(* CODESYS project Visualization.vis.xml

Project tree, tasks and I/O mapping:
  visualisation Visualization
*)

// /Visualization
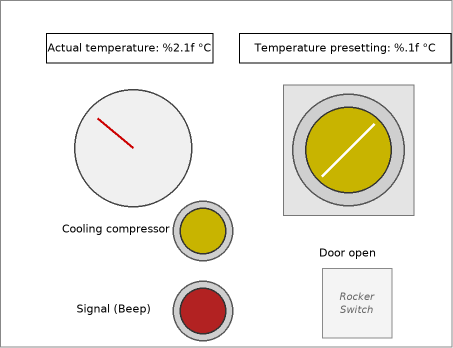
VISUALIZATION Visualization  // 453x348
    Rectangle (46,33 167x30), "Actual temperature: %2.1f °C", text variable: Glob_Var.TempActual
    Lamp1 (168,196 70x70), variable: Glob_Var.Compressor, style: Lamp-Lamp1-Yellow
    Rectangle (239,33 212x30), "Temperature presetting: %.1f °C", text variable: Glob_Var.TempSet
        OnMouseDown: write the text variable via Default, min 3, max 12
    Potentiometer360 (283,84 131x132), variable: Glob_Var.TempSet, style: Potentiometer-Potentiometer360-Yellow, scale format: %.0f, scale 3..13
        p2431819421: Outside
        p518627256: °C
    Meter180 (49,89 168x118), value: Glob_Var.TempActual, style: Meter-Meter180-Gray, scale format: %.1f, scale 0..20
    Rectangle (41,214 150x30), "Cooling compressor"
    Lamp1 (168,276 70x70), variable: Glob_Var.Signal, style: Lamp-Lamp1-Red
    Rectangle (39,294 150x30), "Signal (Beep)"
    RockerSwitch (322,268 70x70), variable: Glob_Var.DoorOpen, behaviour: TOGGLE, style: Switch-RockerSwitch-Gray
    Rectangle (313,238 69x30), "Door open", text variable: Glob_Var.TempSet
END_VISUALIZATION
